// TIA Portal V21 export
// export: Created 2026-10-23T20:42:50.7852386Z, ExportSetting WithDefaults, DisplayName Totally Integrated Automation Portal, DisplayVersion V21 Update 1, DisplayName SINAMICS Startdrive Advanced, DisplayVersion V21 HF2, DisplayName SINAMICS Startdrive G110M, G120, G120C, G120D, G120P, G115D, DisplayVersion V21 HF2, DisplayName SINAMICS Startdrive G130, G150, S120, S150, G200, G220, S200, S210, S220, Innomotics MVD, DisplayVersion V21 HF2, DisplayName STEP 7 Professional, DisplayVersion V21 Update 1, DisplayName STEP 7 Safety, DisplayVersion V21, DisplayName Tech WebApplication, DisplayVersion V21, DisplayName WinCC Basic/Comfort/Advanced, DisplayVersion V21 Update 1, DisplayName WinCC Unified, DisplayVersion V21 Update 1
DATA_BLOCK "DB_Machine"   // DB1
TITLE = Maschinendaten / Machine data
{ S7_Optimized_Access := 'TRUE' }
VERSION : 0.1
// Zentrale Daten der Abfüllmaschine / Central data of the filling machine
// stored: AutoNumber true, DBAccessibleFromOPCUA true, DBAccessibleFromWebserver true, IsOnlyStoredInLoadMemory false, IsRetainMemResEnabled false, IsWriteProtectedInAS false, MemoryReserve 100
   VAR
      MachineOn : Bool := FALSE;   // Maschine eingeschaltet / Machine switched on
      StatusByte : Byte := 16#0F;   // Statusbits als Byte / Status bits as byte
      StatusWord : Word := 16#00FF;   // Statusbits als Wort / Status bits as word
      StatusDWord : DWord := 16#0000_FFFF;   // Statusbits als Doppelwort / Status bits as double word
      StatusLWord : LWord := 16#0000_0000_FFFF_FFFF;   // Statusbits als Langwort / Status bits as long word
      SmallSigned : SInt := -5;   // Kleiner Wert mit Vorzeichen / Small signed value
      SmallUnsigned : USInt := 200;   // Kleiner Wert ohne Vorzeichen / Small unsigned value
      PieceCount : Int := 0;   // Stückzähler mit Vorzeichen / Signed piece counter
      PieceCountUnsigned : UInt := 100;   // Stückzähler ohne Vorzeichen / Unsigned piece counter
      TotalCount : DInt := 0;   // Gesamtzahl der Flaschen / Total number of bottles
      TotalCountUnsigned : UDInt := 0;   // Gesamtzahl der Deckel / Total number of caps
      LongCount : LInt := 0;   // Langer Zähler mit Vorzeichen / Long signed counter
      LongCountUnsigned : ULInt := 0;   // Langer Zähler ohne Vorzeichen / Long unsigned counter
      Temperature : Real := 21.5;   // Produkttemperatur in Grad Celsius / Product temperature in degrees Celsius
      Pressure : LReal := 1.013;   // Leitungsdruck in bar / Line pressure in bar
      CycleTime : Time := T#2S;   // Maschinentaktzeit / Machine cycle time
      PreciseTime : LTime := LT#500US;   // Genaue Taktzeit / Precise cycle time
      LegacyTime : S5Time := S5T#10S;   // Alter Zeitwert / Legacy time value
      ProductionDate : Date := D#2026-01-01;   // Produktionsdatum / Production date
      ShiftStart : Time_Of_Day := TOD#06:00:00;   // Schichtbeginn / Start of the shift
      PreciseShiftStart : LTime_Of_Day := LTOD#06:00:00.000000001;   // Genauer Schichtbeginn / Precise start of the shift
      LegacyTimestamp : Date_And_Time := DT#2026-01-01-06:00:00;   // Alter Zeitstempel / Legacy time stamp
      PreciseTimestamp : LDT := LDT#2026-01-01-06:00:00;   // Genauer Zeitstempel / Precise time stamp
      Separator : Char := 'A';   // Trennzeichen / Separator character
      Symbol : WChar := WCHAR#'B';   // Unicode-Symbol / Unicode symbol
      MachineName : String[20] := 'Filler';   // Maschinenname / Machine name
      OperatorText : WString := WSTRING#'Ready';   // Text für den Bediener / Text for the operator
      LastStart : DTL := DTL#2026-01-01-00:00:00;   // Zeitpunkt des letzten Starts / Time of the last start
      Limits : Struct   // Prozessgrenzen / Process limits
         Minimum : Real := 0.0;   // Untere Grenze / Lower limit
         Maximum : Real := 100.0;   // Obere Grenze / Upper limit
      END_STRUCT;
      Speeds : Array[0..4] of Int;   // Drehzahlstufen / Speed steps
      MainMotor { S7_SetPoint := 'True'} : "UDT_Motor";   // Hauptantrieb / Main drive
      SpeedSetpoint { S7_SetPoint := 'True'} : Real := 50.0;   // Drehzahlsollwert in Prozent / Speed setpoint in percent
      InternalState { ExternalAccessible := 'False'; ExternalVisible := 'False'; ExternalWritable := 'False'} : Int := 0;   // Interner Zustand, für HMI und OPC UA verborgen / Internal state, hidden from HMI and OPC UA
      ReadOnlyValue { ExternalWritable := 'False'} : Real := 0.0;   // Sichtbar, aber von HMI und OPC UA nicht beschreibbar / Visible but not writable from HMI and OPC UA
   END_VAR
   VAR RETAIN
      OperatingHours : DInt := 0;   // Betriebsstunden, remanent / Operating hours, retentive
      RetainedRecipe : Int := 1;   // Last recipe, retentive
   END_VAR
BEGIN
   Speeds[0] := 0;
   Speeds[1] := 10;
   Speeds[2] := 20;
   Speeds[3] := 30;
   Speeds[4] := 40;
END_DATA_BLOCK
